Staubli VAL3: getPointSize.pgx

public program getPointSize(string x_sKey, num& x_nSize)
begin
  x_nSize=size(trajTemp:tTrajItem[x_sKey].pPointItem)
end
